TYPE LaserScan :
STRUCT
	sequence : UDINT;
	startTimestampInNs : ULINT;
	scanDurationInS : REAL;
	angleMinInRad : REAL;
	angleIncrementInRad : REAL;
	count : UINT;
	rangesInM : ARRAY[0..Constants.MAX_SCAN_POINTS - 1] OF REAL;
END_STRUCT
END_TYPE

(* stored: Version 1.1.0.1, ProductVersion 3.1.4026.12
   DUT LaserScan: Id {6202e74c-5eb0-5f6d-bb19-ff61a4ae52c7} *)
